(* IEC 61131-3 sources: PLC_Gen_Frame/Agents4PLC_release/results/task_1778469957, 1 file *)

(* ---- output.ST ---- *)
FUNCTION_BLOCK BakeryOvenControl
VAR_INPUT
    TemperatureSensor : REAL;
    HumiditySensor : REAL;
END_VAR
VAR_OUTPUT
    HeatingElement : BOOL;
    CoolingElement : BOOL;
    HumidityControl : BOOL;
    DehumidityControl : BOOL;
END_VAR

// Generated by DummyPLCGenerator

END_FUNCTION_BLOCK
